DATA_BLOCK "naut_SfcQualifiers_DB"
{ S7_Optimized_Access := 'TRUE' }
VERSION : 0.1
"naut_SfcQualifiers"

BEGIN

END_DATA_BLOCK
